(* IEC 61131-3 sources: rules_plc/examples/external_c_library, 2 files *)

(* ---- fast_math.st ---- *)
{external}
FUNCTION fast_double : DINT
    VAR_INPUT
        x : DINT;
    END_VAR
END_FUNCTION

{external}
FUNCTION fast_negate : DINT
    VAR_INPUT
        x : DINT;
    END_VAR
END_FUNCTION

(* A stateful {external} FUNCTION_BLOCK, unlike fast_double/fast_negate above
-- exercises the same weak-stub mechanism for the struct-plus-function ABI
FUNCTION_BLOCK compiles to, rather than a plain value-returning function.
    *)
    {external}
    FUNCTION_BLOCK fast_counter
        VAR_INPUT
            step : DINT;
        END_VAR
        VAR
            state: DINT;
        END_VAR
        VAR_OUTPUT
            value : DINT;
        END_VAR
    END_FUNCTION_BLOCK

(* ---- fast_math_bin.st ---- *)
PROGRAM fast_math_bin
    VAR
        a : REAL := 12.5;
        b : REAL := 3.5;
        sum : REAL;
        diff : REAL;
        prod : REAL;
        quot : REAL;
        valid_div : BOOL;
    END_VAR

    sum := a + b;
    diff := a - b;
    prod := a * b;

    valid_div := b <> 0.0;
    IF valid_div THEN
        quot := a / b;
    ELSE
        quot := 0.0;
    END_IF;

END_PROGRAM
